(*
    Command and status view of a pneumatic actuator. Insert() and Retract() raise
    the same requests as the CMD:IN and CMD:OUT PVs. Both requests together cancel
    each other.
*)
INTERFACE I_PneumaticActuator

METHOD Insert
VAR_INPUT
END_VAR
END_METHOD

METHOD Retract
VAR_INPUT
END_VAR
END_METHOD

PROPERTY Busy : BOOL
GET
END_GET
END_PROPERTY

PROPERTY Done : BOOL
GET
END_GET
END_PROPERTY

PROPERTY Error : BOOL
GET
END_GET
END_PROPERTY

PROPERTY MpsOk : BOOL
GET
END_GET
END_PROPERTY

PROPERTY State : E_PnuematicActuatorPositionState
GET
END_GET
END_PROPERTY

END_INTERFACE

(* stored: Version 1.1.0.1
   Itf I_PneumaticActuator: Id {a3f0aa9b-1939-4de3-ba56-c149a572d90a}
   Method Insert: Id {629b967c-f1f3-4e00-ac8f-3a6e29974957}
   Method Retract: Id {6ac4bc52-d297-4926-b458-b138f94e3b88}
   Property Busy: Id {b5a7dc1a-8b3f-4753-baaa-de7326ca7b6f}
   Get Get: Id {4260e850-c541-415e-a638-c0d93ecc4bf6}
   Property Done: Id {0adecd69-56be-46c0-aea1-10ef7fc17842}
   Get Get: Id {fdaa5543-3d3a-4379-9dc6-ee5513fbf77e}
   Property Error: Id {04f99924-35cd-4b63-b17d-191e9263ed83}
   Get Get: Id {e18ab759-bd4b-4b69-a635-99fd0eff6522}
   Property MpsOk: Id {de9e9118-a3bc-4fa6-b14d-4c7b193413e2}
   Get Get: Id {c645692a-4000-41f4-979b-f0b7a7a88447}
   Property State: Id {c3e5c914-d8c8-4134-8136-5bdc5bbac04e}
   Get Get: Id {3236e6cc-c340-4964-a321-379ad397b454} *)
